  global target_g_table = [
  	"NaCl", "spatula_L", "6.5",
  	"NaCl", "spatula_M", "1.5",
  	"NaCl", "spatula_S", "0.135",

  	"Mannitol", "spatula_L", "2.85",
  	"Mannitol", "spatula_M", "0.8",
  	"Mannitol", "spatula_S", "0.075",

  	"CCS", "spatula_L", "2.45",
  	"CCS", "spatula_M", "0.6",
  	"CCS", "spatula_S", "0.075",

  	"lactose_loose", "spatula_L", "1.6",
  	"lactose_loose", "spatula_M", "0.5",
  	"lactose_loose", "spatula_S", "0.05",

  	"Magnesium_sterate", "spatula_flat_M", "0.6",
  	"Magnesium_sterate", "spatula_flat_S", "0.25",

  	"lactose_fine", "spatula_flat_M", "1.0",
  	"lactose_fine", "spatula_flat_S", "0.5"]

  def get_target_g(Pow_name, spat_name):
  	local i = 0
  	local n = length(target_g_table)
  	while (i < n):
  		if (target_g_table[i] == Pow_name and target_g_table[i+1] == spat_name):
  			return to_num(target_g_table[i+2])
  		end
  		i = i+3
  	end
  	popup("No target_g match for: ", Pow_name, ", ", spatula)

  end
  def auto_tilt_and_scoop(W_now, target_weight, Weight_value):
  	level = compute_level_percent(W_now, Weight_value)

  	#global angle_deg = compute_tilt_deg(level)

  	#if(level>=10.0):
  		#target_g = 2.850
  	#elif(level<10.0 and level >=1.0):
  		#target_g= 0.8
  	#else:
  		#target_g = 0.060
  	#end


  	#if (Task =="Emptying"):
  		#if (level>10.0):
  			#target_g = 2.850
  		#elif (level<=10.0 and level >1.0):
  			#target_g = 0.8
  		#else:
  			#target_g = 0.060
  		#end
  	#elif (Task == "Dosing"):
  		#if (level>10.0 and diff>=3.5):
  			#target_g = 2.85
  		#elif (level>10.0 and diff<3.5):
  			#target_g = 0.8
  		#elif (level<=10.0 and level >1.0):
  			#target_g = 0.8
  		#else:
  			#target_g = 0.06
  		#end
  	#end

  	global spatula = select_spatula(Pow_name, level, diff)
  	global target_g = get_target_g(Pow_name, spatula)

  	global scoop_depth = compute_scoop_depth(level, Weight_value, target_g)

  	tilt(level)
  	#P_center = get_actual_tcp_pose()

  	if (scoop_ct < 5 and g_prev_cum_w>0.0):
  		#local scoop_g = scoop_g
  		local error = target_g - scoop_g
  		error_sum = error_sum + error
  		error_sq_sum = error_sq_sum + error*error
  		scoop_ct = scoop_ct+1

  		if (scoop_ct==5):
  			local avg_error = error_sum/5.0
  			#local std_dev = sqrt(error_sq_sum/5.0) - (avg_error*avg_error))

  			if (my_abs(avg_error)>1.0):
  				g_k = 0.055
  				g_alpha = 0.85
  			elif (my_abs(avg_error)>0.6):
  				g_k= 0.045
  				g_alpha =0.75
  			elif (my_abs(avg_error)> 0.3):
  				g_k = 0.035
  				g_alpha = 0.65
  			elif (my_abs(avg_error)>0.1):
  				g_k = 0.025
  				g_alpha = 0.55
  			else:
  				g_k = 0.015
  				g_alpha = 0.45
  			end
  		end
  	end

  	scoop_powder(P_center)
  end


  def after_scoop():
  	tilt_send(angle_deg)
  	sleep(0.5)
  	movel(lifted_pose, a=0.05, v=0.2)
  	movel(tilted_pose_in_base, a=0.05, v=0.2)
  	set_analog_out(0,0.4)
  	movel(pose_trans(tilted_pose_in_base, p[-0.01,0,0,0,0,2.0]), a=0.05, v=0.2)
  	set_analog_out(0,0.0)
  	movel(lifted_pose, a=0.05, v=0.2)
  	tilt_to_home()
  end
  $ 23 "Script: Weight_scale_socket.script"
  def get_weight():
  	socket_open("192.168.12.190", 3002)
  	sleep(0.2)
  	textmsg("socket opened successfully!")
  	socket_send_string("GET_WEIGHT")
  	sync()
  	sleep(0.5)
  	receiveFromServ = socket_read_ascii_float(6)
  	while (receiveFromServ[0] <1):
  		sleep(0.5)
  		receiveFromServ = socket_read_ascii_float(1)
  		textmsg("retrying read:", receiveFromServ)
  	end
  	textmsg("Received weight:", receiveFromServ[1])
  	socket_close()
  	sleep(0.2)
  	return receiveFromServ[1]
  end

  def tare_scale():
  	socket_open("192.168.12.190", 3002)
  	socket_send_string("TARE")
  	sleep(0.5)
  	socket_close()
  end

  def zero_scale():
  	socket_open("192.168.12.190", 3002)
  	socket_send_string("ZERO")
  	sleep(0.5)
  	socket_close()
  end

  def log_weight():
  	socket_open("192.168.12.190", 3002)
  	socket_send_string("LOG_WEIGHT")
  	sleep(0.5)
  	socket_close()
  end
  $ 24 "BeforeStarts"
  $ 25 "uLM"
  $ 26 "CMD_Stop≔ False "
  global CMD_Stop=  False
  $ 27 "CMD_Abort≔ False "
  global CMD_Abort=  False
  $ 28 "CMD_Clear≔ False "
  global CMD_Clear=  False
  $ 29 "STATE≔1"
  global STATE=1
  $ 30 "STATE_Info≔''"
  global STATE_Info=""
  $ 31 "ARM_Referenced≔ False "
  global ARM_Referenced=  False
  $ 32 "zero_ftsensor()"
  zero_ftsensor()
  $ 33 "poses init"
  $ 34 "PSE_A≔p[0,0,0,0,0,0]"
  global PSE_A=p[0,0,0,0,0,0]
  $ 35 "PSE_A_H≔p[0,0,0,0,0,0]"
  global PSE_A_H=p[0,0,0,0,0,0]
  $ 36 "PSE_R≔p[0,0,0,0,0,0]"
  global PSE_R=p[0,0,0,0,0,0]
  $ 37 "PSE_R_H≔p[0,0,0,0,0,0]"
  global PSE_R_H=p[0,0,0,0,0,0]
  $ 38 "PSE_T≔p[0,0,0,0,0,0]"
  global PSE_T=p[0,0,0,0,0,0]
  $ 39 "PSE_T_H≔p[0,0,0,0,0,0]"
  global PSE_T_H=p[0,0,0,0,0,0]
  $ 40 "PSE_C_E≔p[0,0,0,0,0,0]"
  global PSE_C_E=p[0,0,0,0,0,0]
  $ 41 "PSE_C_H≔p[0,0,0,0,0,0]"
  global PSE_C_H=p[0,0,0,0,0,0]
  $ 42 "PSE_C_S≔p[0,0,0,0,0,0]"
  global PSE_C_S=p[0,0,0,0,0,0]
  $ 43 "init_home_by_cartesian_pose(p[0,-0.400,0.300,0,0,0])"
  init_home_by_cartesian_pose(p[0,-0.400,0.300,0,0,0])
  $ 44 "Clearing"
  $ 45 "reset_error()"
  reset_error()
  $ 46 "reset_warning()"
  reset_warning()
  $ 47 "uGo"
  $ 49 "ugo_init( True ,'http://192.168.12.120:10001')"
  ugo_init(  True  ,"http://192.168.12.120:10001")
  $ 50 "ugo_update_outputs()"
  ugo_update_outputs()
  $ 51 "App"
  $ 52 "'ADD APPLICATION SPECIFIC COMMANDS'"
  # 'ADD APPLICATION SPECIFIC COMMANDS'
  $ 53 "Tools"
  $ 54 "OBJ_Picked≔gripper_has_object()"
  global OBJ_Picked=gripper_has_object()
  $ 55 "If OBJ_Picked"
  if (OBJ_Picked):
    # begin: URCap Program Node
    #   Source: Robotiq_Grippers, 1.8.4.4844, Robotiq Inc.
    #   Type: Gripper Activate
    $ 56 "Gripper Activate"

    kill rq_gripper_communication_thread
    rq_gripper_communication_thread_started = False

    rq_init_comm_if_connected(9, "1")
    rq_init_comm_if_connected(2, "2")
    rq_init_comm_if_connected(3, "3")
    rq_init_comm_if_connected(4, "4")
    rq_print_connected_grippers()
    rq_gripper_communication_thread = run rq_gripper_communication()

    while(not rq_gripper_communication_thread_started):
        sync()
    end

    rq_set_max_current_for_all_grippers()

    reset_and_activate = False

    rq_activate_all_grippers(False)
    # end: URCap Program Node
  else:
    $ 57 "Else" "noBreak"
    # begin: URCap Program Node
    #   Source: Robotiq_Grippers, 1.8.4.4844, Robotiq Inc.
    #   Type: Gripper Activate
    $ 58 "Gripper Reset and Activate"

    kill rq_gripper_communication_thread
    rq_gripper_communication_thread_started = False

    rq_init_comm_if_connected(9, "1")
    rq_init_comm_if_connected(2, "2")
    rq_init_comm_if_connected(3, "3")
    rq_init_comm_if_connected(4, "4")
    rq_print_connected_grippers()
    rq_gripper_communication_thread = run rq_gripper_communication()

    while(not rq_gripper_communication_thread_started):
        sync()
    end

    rq_set_max_current_for_all_grippers()

    reset_and_activate = True

    rq_activate_all_grippers(True)
    # end: URCap Program Node
  end
  $ 59 "zero_ftsensor()"
  zero_ftsensor()
  $ 60 "EXTT"
  $ 61 "Set GRP_3F_Enable=Off"
  set_standard_digital_out(4, False)
  $ 62 "Set DO[6]=Off"
  set_standard_digital_out(6, False)
  $ 63 "Set GRP_3F_Decap=Off"
  set_standard_digital_out(3, False)
  $ 64 "Set GRP_3F_Cap=Off"
  set_standard_digital_out(2, False)
  $ 65 "Set GRP_3F_Open=Off"
  set_standard_digital_out(5, False)
  $ 66 "PSE_T≔get_tool_free_pose(dir=[0,0,0.150], move_in_base_frame=True)"
  global PSE_T=get_tool_free_pose(dir=[0,0,0.150], move_in_base_frame=True)
  $ 67 "If is_reachable(Base_const, [PSE_T])"
  if (is_reachable(p[0.0,0.0,0.0,0.0,0.0,0.0], [PSE_T])):
    $ 68 "MoveL"
    $ 69 "PSE_T" "breakAfter"
    movel(PSE_T, a=1.2, v=0.15)
  end
  $ 70 "powder dispensing variable init"
  $ 71 "Start_thread≔ False "
  global Start_thread=  False
  $ 72 "vib_mot_thread≔ False "
  global vib_mot_thread=  False
  $ 73 "kp≔0.0005"
  global kp=0.0005
  $ 74 "ki≔0.005"
  global ki=0.005
  $ 75 "kd≔0.02"
  global kd=0.02
  $ 76 "dt≔0.02"
  global dt=0.02
  $ 77 "Integral_error≔0"
  global Integral_error=0
  $ 78 "current_error≔0"
  global current_error=0
  $ 79 "previous_error≔0"
  global previous_error=0
  $ 80 "tilt_increment≔0"
  global tilt_increment=0
  $ 81 "tilt_angle≔0"
  global tilt_angle=0
  $ 82 "diff≔0"
  global diff=0
  $ 83 "current_pose≔get_actual_tcp_pose()"
  global current_pose= get_actual_tcp_pose ()
  $ 84 "Relative_trans≔p[0, 0, -0.035, 0, 0, 0]"
  global Relative_trans=p[0, 0, -0.035, 0, 0, 0]
  $ 85 "ContA_plc_offst≔p[-0.00205, 0.02547, 0.03730, -0.03, -2.183, 6.165]"
  global ContA_plc_offst=p[-0.00205, 0.02547, 0.03730, -0.03, -2.183, 6.165]
  $ 86 "PowA_50_offset≔p[0.21808, -0.19943, 0.06584, 0, 0, 0]"
  global PowA_50_offset=p[0.21808, -0.19943, 0.06584, 0, 0, 0]
  $ 88 "tilt_init_reference()"
  tilt_init_reference()
  $ 89 "switch_spat_M≔ True "
  global switch_spat_M=  True
  $ 90 "switch_spat_S≔ True "
  global switch_spat_S=  True
  $ 698 "Thread_1"
  thread Thread_1():
    while (True):
      $ 699 "If Start_thread≟ True "
      if (Start_thread ==   True  ):
        $ 700 "Weight_value≔get_weight()"
        global Weight_value=get_weight()
        $ 701 "Wait: 0.1"
        sleep(0.1)
        $ 702 "sync()"
        sync()
      end
    end
  end
  threadId_Thread_1 = run Thread_1()
  while (True):
    $ 91 "Robot Program"
    $ 92 "MAIN"
    $ 93 "command_manager(external_control='uGO', cond_suspend=(ITM_Manipulated and AMR_AtTarget and AMR_Charging and AMR_Battery<40), cond_unsuspend=(AMR_Battery≟60))"
    command_manager(external_control="uGO", cond_suspend=(ITM_Manipulated  and  AMR_AtTarget  and  AMR_Charging  and  AMR_Battery<40), cond_unsuspend=(AMR_Battery == 60))
    $ 94 "log_state(STATE_Info)"
    log_state(STATE_Info)
    $ 95 "Switch STATE"
    switch_1 = STATE
    $ 96 "Case 1"
    if (1 == switch_1):
      $ 97 "Stopping"
      $ 98 "STATE_Info≔'Stopping'"
      global STATE_Info="Stopping"
      $ 99 "end_freedrive_mode()"
      end_freedrive_mode()
      $ 100 "Set"
      set_tcp(p[0.0,0.0,0.161,3.1415,0.0,0.0])
      $ 101 "PSE_T≔get_tool_free_pose(dir=[0,0,0.150], move_in_base_frame=True)"
      global PSE_T=get_tool_free_pose(dir=[0,0,0.150], move_in_base_frame=True)
      $ 102 "If is_reachable(Base_const, [PSE_T])"
      if (is_reachable(p[0.0,0.0,0.0,0.0,0.0,0.0], [PSE_T])):
        $ 103 "MoveL"
        $ 104 "PSE_T" "breakAfter"
        movel(PSE_T, a=1.2, v=0.15)
      end
      $ 105 "do_transition(keep_rxry=OBJ_Picked, r=0)"
      do_transition(keep_rxry=OBJ_Picked, r=0)
      $ 115 "If stopping() and AMR_Done"
      if (stopping()  and  AMR_Done):
        $ 116 "STATE≔2"
        global STATE=2
        $ 117 "ugo_update_outputs()"
        ugo_update_outputs()
      end
    elif (2 == switch_1):
      $ 118 "Case 2"
      $ 119 "Stopped"
      $ 120 "STATE_Info≔'Stopped'"
      global STATE_Info="Stopped"
      $ 122 "If CMD_Reset"
      if (CMD_Reset):
        $ 123 "STATE≔3"
        global STATE=3
        $ 124 "ugo_update_outputs()"
        ugo_update_outputs()
      end
    elif (3 == switch_1):
      $ 125 "Case 3"
      $ 126 " Resetting"
      $ 127 "STATE_Info≔'Resetting'"
      global STATE_Info="Resetting"
      $ 128 "uML"
      $ 129 "reset_error()"
      reset_error()
      $ 130 "reset_warning()"
      reset_warning()
      $ 131 "PROCESS_Step≔0"
      global PROCESS_Step=0
      $ 132 "PROCESS_Info≔''"
      global PROCESS_Info=""
      $ 133 "ARM_Referenced≔ False "
      global ARM_Referenced=  False
      $ 134 "WRK_Done≔ False "
      global WRK_Done=  False
      $ 135 "ITM_Prepared≔ False "
      global ITM_Prepared=  False
      $ 136 "ITM_Manipulated≔ False "
      global ITM_Manipulated=  False
      $ 137 "STP≔0"
      global STP=0
      $ 138 "Action≔0"
      global Action=0
      $ 139 "Action_Info≔''"
      global Action_Info=""
      $ 140 "ITM_ID≔0"
      global ITM_ID=0
      $ 141 "JIG≔0"
      global JIG=0
      $ 142 "JIG_Slot≔0"
      global JIG_Slot=0
      $ 143 "Task_info≔''"
      global Task_info=""
      $ 144 "Set"
      set_tcp(p[0.0,0.0,0.161,3.1415,0.0,0.0])
      $ 145 "App"
      $ 146 "'ADD APPLICATION SPECIFIC COMMANDS'"
      # 'ADD APPLICATION SPECIFIC COMMANDS'
      $ 147 "OBJ_Type≔0"
      global OBJ_Type=0
      $ 148 "OBJ_Nbr≔0"
      global OBJ_Nbr=0
      $ 149 "If CNT_Rack_Output≥50"
      if (CNT_Rack_Output >= 50):
        $ 150 "CNT_Rack_Output≔0"
        global CNT_Rack_Output=0
      end
      $ 151 "TASK≔struct(ID=0, NAVI=struct(target=0, footprint=0, protectiveOff=0, dock=0), WORK=struct(ITM_ID_Src=0, JIG_ID_Src=0, OBJ_Nbr_Src=0, ACT_Src=0, ITM_ID_Tgt=0, JIG_ID_Tgt=0, OBJ_Nbr_Tgt=0, ACT_Tgt=0, OBJ_Type=0))"
      global TASK=struct(ID=0, NAVI=struct(target=0, footprint=0, protectiveOff=0, dock=0), WORK=struct(ITM_ID_Src=0, JIG_ID_Src=0, OBJ_Nbr_Src=0, ACT_Src=0, ITM_ID_Tgt=0, JIG_ID_Tgt=0, OBJ_Nbr_Tgt=0, ACT_Tgt=0, OBJ_Type=0))
      $ 153 "If resetting() and AMR_Done"
      if (resetting()  and  AMR_Done):
        $ 154 "STATE≔4"
        global STATE=4
        $ 155 "ugo_update_outputs()"
        ugo_update_outputs()
      end
    elif (4 == switch_1):
      $ 156 "Case 4"
      $ 157 "Idle"
      $ 158 "STATE_Info≔'Idle'"
      global STATE_Info="Idle"
      $ 159 "If CMD_Start"
      if (CMD_Start):
        $ 160 "STATE≔5"
        global STATE=5
        $ 161 "ugo_update_outputs()"
        ugo_update_outputs()
      end
    elif (5 == switch_1):
      $ 162 "Case 5"
      $ 163 "Starting"
      $ 164 "STATE_Info≔'Starting'"
      global STATE_Info="Starting"
      $ 165 "'ADD COMMANDS WHAT TO START WITH'"
      # 'ADD COMMANDS WHAT TO START WITH'
      $ 167 "get ugo data"
      $ 168 "Assign Tasks"
      $ 169 "TASK.ID = ugo_get_task()"
      TASK.ID = ugo_get_task()
      $ 170 "If TASK.ID≟1"
      if (TASK.ID == 1):
        $ 171 "Task_info≔'Charge'"
        global Task_info="Charge"
        $ 172 "Parameters"
        $ 173 "AMR_PosTarget≔1"
        global AMR_PosTarget=1
      else:
        $ 174 "ElseIf TASK.ID≟9"
        if (TASK.ID == 9):
          $ 175 "'Pick Sarstedt Rack from Variable source'"
          # 'Pick Sarstedt Rack from Variable source'
          $ 176 "Task_info≔'Navigate to Target'"
          global Task_info="Navigate to Target"
          $ 177 "Parameters"
          $ 178 "AMR_PosTarget≔UGO.read_input('00','ITM_ID')"
          global AMR_PosTarget=UGO.read_input("00","ITM_ID")
        else:
          $ 179 "ElseIf TASK.ID≟49"
          if (TASK.ID == 49):
            $ 180 "Task_info≔'Pick Containers'"
            global Task_info="Pick Containers"
            $ 181 "Parameters"
            $ 182 "ITM_ID≔1"
            global ITM_ID=1
            $ 183 "OBJ_Type≔6"
            global OBJ_Type=6
            $ 184 "JIG≔15"
            global JIG=15
            $ 185 "AMR_PosTarget≔3"
            global AMR_PosTarget=3
          else:
            $ 186 "ElseIf TASK.ID≟50"
            if (TASK.ID == 50):
              $ 187 "Task_info≔'Decap Containers'"
              global Task_info="Decap Containers"
              $ 188 "Parameters"
              $ 189 "ITM_ID≔1"
              global ITM_ID=1
              $ 190 "OBJ_Type≔6"
              global OBJ_Type=6
              $ 191 "JIG≔16"
              global JIG=16
              $ 192 "AMR_PosTarget≔5"
              global AMR_PosTarget=5
            else:
              $ 193 "ElseIf TASK.ID≟51"
              if (TASK.ID == 51):
                $ 194 "Task_info≔'Detect Spatula and transfer powder'"
                global Task_info="Detect Spatula and transfer powder"
                $ 195 "Parameters"
                $ 196 "ITM_ID≔1"
                global ITM_ID=1
                $ 197 "Target_weight≔(UGO.read_input('00','Target_weight'))/1000"
                global Target_weight=(UGO.read_input("00","Target_weight"))/1000
                $ 198 "OBJ_Type≔8"
                global OBJ_Type=8
                $ 199 "JIG≔16"
                global JIG=16
                $ 200 "AMR_PosTarget≔5"
                global AMR_PosTarget=5
              else:
                $ 201 "ElseIf TASK.ID≟52"
                if (TASK.ID == 52):
                  $ 202 "Task_info≔'Pick PowderA'"
                  global Task_info="Pick PowderA"
                  $ 203 "Parameters"
                  $ 204 "ITM_ID≔1"
                  global ITM_ID=1
                  $ 205 "OBJ_Type≔6"
                  global OBJ_Type=6
                  $ 206 "JIG≔15"
                  global JIG=15
                  $ 207 "AMR_PosTarget≔3"
                  global AMR_PosTarget=3
                else:
                  $ 208 "ElseIf TASK.ID≟53"
                  if (TASK.ID == 53):
                    $ 209 "Task_info≔'Decap PowderA'"
                    global Task_info="Decap PowderA"
                    $ 210 "Parameters"
                    $ 211 "ITM_ID≔1"
                    global ITM_ID=1
                    $ 212 "OBJ_Type≔6"
                    global OBJ_Type=6
                    $ 213 "JIG≔1"
                    global JIG=1
                    $ 214 "AMR_PosTarget≔5"
                    global AMR_PosTarget=5
                  else:
                    $ 215 "ElseIf TASK.ID≟54"
                    if (TASK.ID == 54):
                      $ 216 "Task_info≔'Empty PowderA'"
                      global Task_info="Empty PowderA"
                      $ 217 "Parameters"
                      $ 218 "ITM_ID≔1"
                      global ITM_ID=1
                      $ 219 "Target_weight≔(UGO.read_input('00','Target_weight'))/1000"
                      global Target_weight=(UGO.read_input("00","Target_weight"))/1000
                      $ 220 "W_now≔(UGO.read_input('00','Container_weight'))/1000"
                      global W_now=(UGO.read_input("00","Container_weight"))/1000
                      $ 221 "Powder_name≔(UGO.read_input('00','Powder_name'))"
                      global Powder_name=(UGO.read_input("00","Powder_name"))
                      $ 222 "OBJ_Type≔6"
                      global OBJ_Type=6
                      $ 223 "JIG≔17"
                      global JIG=17
                      $ 224 "AMR_PosTarget≔5"
                      global AMR_PosTarget=5
                    else:
                      $ 225 "ElseIf TASK.ID≟55"
                      if (TASK.ID == 55):
                        $ 226 "Task_info≔'Place PowderA'"
                        global Task_info="Place PowderA"
                        $ 227 "Parameters"
                        $ 228 "ITM_ID≔1"
                        global ITM_ID=1
                        $ 229 "OBJ_Type≔6"
                        global OBJ_Type=6
                        $ 230 "JIG≔21"
                        global JIG=21
                        $ 231 "AMR_PosTarget≔5"
                        global AMR_PosTarget=5
                      else:
                        $ 232 "ElseIf TASK.ID≟56"
                        if (TASK.ID == 56):
                          $ 233 "Task_info≔'Dose Powder'"
                          global Task_info="Dose Powder"
                          $ 234 "Parameters"
                          $ 235 "ITM_ID≔1"
                          global ITM_ID=1
                          $ 236 "Target_weight≔(UGO.read_input('00','Target_weight'))/1000"
                          global Target_weight=(UGO.read_input("00","Target_weight"))/1000
                          $ 237 "W_now≔(UGO.read_input('00','Container_weight'))/1000"
                          global W_now=(UGO.read_input("00","Container_weight"))/1000
                          $ 238 "Pow_name≔(UGO.read_input('00','Powder_name'))"
                          global Pow_name=(UGO.read_input("00","Powder_name"))
                          $ 239 "OBJ_Type≔6"
                          global OBJ_Type=6
                          $ 240 "JIG≔17"
                          global JIG=17
                          $ 241 "AMR_PosTarget≔5"
                          global AMR_PosTarget=5
                        else:
                          $ 242 "Else" "noBreak"
                          $ 243 "set_error(ERROR_WRONG_ORDER)"
                          set_error(ERROR_WRONG_ORDER)
                        end
                      end
                    end
                  end
                end
              end
            end
          end
        end
      end
      $ 244 "test ugo"
      $ 245 "Wait: 0.2"
      sleep(0.2)
      $ 246 "ugo_update_outputs()"
      ugo_update_outputs()
      $ 247 "If starting() and AMR_Done"
      if (starting()  and  AMR_Done):
        $ 248 "log_message(Task_info, 'New Task: ')"
        log_message(Task_info, "New Task: ")
        $ 249 "log_message(to_str(TASK.ID), 'Task_ID: ')"
        log_message(to_str(TASK.ID), "Task_ID: ")
        $ 250 "do_transition(keep_rxry=OBJ_Picked)"
        do_transition(keep_rxry=OBJ_Picked)
        $ 251 "STATE≔6"
        global STATE=6
        $ 252 "ugo_update_outputs()"
        ugo_update_outputs()
      end
    elif (6 == switch_1):
      $ 253 "Case 6"
      $ 254 "Execute"
      $ 255 "STATE_Info≔'Execute'"
      global STATE_Info="Execute"
      $ 256 "If  not CMD_Hold and not CMD_Suspend"
      global thread_flag_256=0
      thread Thread_if_256():
        $ 257 "Switch PROCESS_Step"
        switch_2 = PROCESS_Step
        $ 258 "Case 0"
        if (0 == switch_2):
          $ 259 "PROCESS_Info≔'process control'"
          global PROCESS_Info="process control"
          $ 260 "log_process(PROCESS_Info)"
          log_process(PROCESS_Info)
          $ 261 "process control"
          $ 262 "If  not AMR_AtTarget"
          if (  not  AMR_AtTarget):
            $ 263 "PROCESS_Step≔1"
            global PROCESS_Step=1
          else:
            $ 264 "ElseIf (( not ITM_Prepared and  not WRK_Done) or (ITM_Prepared and WRK_Done))"
            if (((  not  ITM_Prepared  and    not  WRK_Done)  or  (ITM_Prepared  and  WRK_Done))):
              $ 265 "PROCESS_Step≔2"
              global PROCESS_Step=2
            else:
              $ 266 "ElseIf  not WRK_Done"
              if (  not  WRK_Done):
                $ 267 "PROCESS_Step≔3"
                global PROCESS_Step=3
              else:
                $ 268 "Else" "noBreak"
                $ 269 "task finished"
                $ 270 "PROCESS_Info≔''"
                global PROCESS_Info=""
                $ 271 "STATE≔7"
                global STATE=7
                $ 272 "ugo_update_outputs()"
                ugo_update_outputs()
              end
            end
          end
        elif (1 == switch_2):
          $ 273 "Case 1"
          $ 274 "navigate"
          $ 275 "'MOVING THE uML'"
          # 'MOVING THE uML'
          $ 276 "PROCESS_Info≔'move to target'"
          global PROCESS_Info="move to target"
          $ 277 "log_process(PROCESS_Info)"
          log_process(PROCESS_Info)
          $ 278 "If TASK.ID≟1"
          if (TASK.ID == 1):
            $ 279 "Action≔51"
            global Action=51
          else:
            $ 280 "Else" "noBreak"
            $ 281 "Action≔52"
            global Action=52
          end
          $ 283 "If AMR_Done"
          if (AMR_Done):
            $ 284 "PROCESS_Step≔0"
            global PROCESS_Step=0
          end
        elif (2 == switch_2):
          $ 285 "Case 2"
          $ 286 "prepare"
          $ 287 "'THINGS THAT HAVE TO BE DONE ONCE IN A SEQUENCE,WORKFLOW'"
          # 'THINGS THAT HAVE TO BE DONE ONCE IN A SEQUENCE,WORKFLOW'
          $ 288 "PROCESS_Info≔'prepare for work'"
          global PROCESS_Info="prepare for work"
          $ 289 "log_process(PROCESS_Info)"
          log_process(PROCESS_Info)
          $ 290 "If TASK.WORK.ITM_ID_Src>1"
          if (TASK.WORK.ITM_ID_Src>1):
            $ 291 "ITM_ID≔TASK.WORK.ITM_ID_Src"
            global ITM_ID=TASK.WORK.ITM_ID_Src
          else:
            $ 292 "ElseIf TASK.WORK.ITM_ID_Tgt>1"
            if (TASK.WORK.ITM_ID_Tgt>1):
              $ 293 "ITM_ID≔TASK.WORK.ITM_ID_Tgt"
              global ITM_ID=TASK.WORK.ITM_ID_Tgt
            end
          end
          $ 294 "If  not ARM_Referenced and (ITM_ID≠0)"
          if (  not  ARM_Referenced  and  (ITM_ID != 0)):
            $ 295 "STP≔1"
            global STP=1
          else:
            $ 296 "ElseIf ARM_Referenced or (ITM_ID≟0)"
            if (ARM_Referenced  or  (ITM_ID == 0)):
              $ 297 "STP≔2"
              global STP=2
            end
          end
          $ 298 "Switch STP"
          switch_3 = STP
          $ 299 "Case 1"
          if (1 == switch_3):
            $ 300 "reference"
            $ 301 "STP_Info≔'reference at target position'"
            global STP_Info="reference at target position"
            $ 302 "log_step(STP_Info)"
            log_step(STP_Info)
            $ 303 "If ITM_ID≟1"
            if (ITM_ID == 1):
              $ 304 "CAM_Done≔ True "
              global CAM_Done=  True
            else:
              $ 305 "Else" "noBreak"
              $ 306 "Action≔131"
              global Action=131
              $ 307 "Call Sub_Vision_V18"
              Sub_Vision_V18()
            end
            $ 309 "If CAM_Done and  not ERROR.FLAG"
            if (CAM_Done  and    not  ERROR.FLAG):
              $ 310 "log_step('ARM referenced')"
              log_step("ARM referenced")
              $ 311 "ARM_Referenced≔ True "
              global ARM_Referenced=  True
            end
          elif (2 == switch_3):
            $ 312 "Case 2"
            $ 313 "manipulate"
            $ 314 "STP_Info≔'manipulate item'"
            global STP_Info="manipulate item"
            $ 315 "log_step(STP_Info)"
            log_step(STP_Info)
            $ 316 "'In case pressing button is needed'"
            # 'In case pressing button is needed'
            $ 317 "If found_in_list(ITM_ID, ITM_ID_List)"
            if (found_in_list(ITM_ID, ITM_ID_List)):
              $ 318 "Switch ITM_ID"
              switch_4 = ITM_ID
              $ 319 "Case 0"
              if (0 == switch_4):
                $ 320 "ITM_Manipulated≔ not ITM_Manipulated"
                global ITM_Manipulated=  not  ITM_Manipulated
              elif (1 == switch_4):
                $ 321 "Case 1"
                $ 322 "ITM_Manipulated≔ not ITM_Manipulated"
                global ITM_Manipulated=  not  ITM_Manipulated
              elif (2 == switch_4):
                $ 323 "Case 2"
              else:
                $ 333 "Default Case"
                $ 334 "ITM_Manipulated≔ not ITM_Manipulated"
                global ITM_Manipulated=  not  ITM_Manipulated
              end
            end
          end
          $ 335 "ITM_Prepared≔(ITM_Manipulated or  not found_in_list(ITM_ID, ITM_ID_List)) and (ARM_Referenced or ITM_ID≟0) and  not WRK_Done"
          global ITM_Prepared=(ITM_Manipulated  or    not  found_in_list(ITM_ID, ITM_ID_List))  and  (ARM_Referenced  or  ITM_ID == 0)  and    not  WRK_Done
          $ 336 "STP≔0"
          global STP=0
          $ 337 "STP_Info≔''"
          global STP_Info=""
          $ 338 "PROCESS_Step≔0"
          global PROCESS_Step=0
        elif (3 == switch_2):
          $ 339 "Case 3"
          $ 340 "work"
          $ 341 "'ADD EVERY MACHINE, OBJECT, STATION TO WORK ON'"
          # 'ADD EVERY MACHINE, OBJECT, STATION TO WORK ON'
          $ 342 "Switch ITM_ID"
          switch_3 = ITM_ID
          $ 343 "Case 1"
          if (1 == switch_3):
            $ 344 "uLM"
            $ 345 "If TASK.ID≟12"
            if (TASK.ID == 12):
              $ 346 "fill racks"
              $ 347 "Action≔151"
              global Action=151
              $ 348 "Call Sub_Vision_V18"
              Sub_Vision_V18()
              $ 349 "If  not ERROR.FLAG"
              if (  not  ERROR.FLAG):
                $ 350 "Actions for the task"
                $ 351 "Action≔1"
                global Action=1
                $ 352 "JIG≔2"
                global JIG=2
                $ 353 "JIG_Slot≔CAM_Result[0]"
                global JIG_Slot=CAM_Result[0]
                $ 354 "OBJ_Nbr≔CAM_Result[0]"
                global OBJ_Nbr=CAM_Result[0]
                $ 355 "OBJ_Type≔2"
                global OBJ_Type=2
                $ 356 "Call Sub_Action_V4"
                Sub_Action_V4()
                $ 357 "If OBJ_Picked"
                if (OBJ_Picked):
                  $ 358 "CAM_Result.remove(0)"
                  CAM_Result.remove(0)
                  $ 359 "PRC_TubCounter≔PRC_TubCounter+1"
                  global PRC_TubCounter=PRC_TubCounter+1
                  $ 360 "If PRC_TubCounter%4≟0"
                  if (PRC_TubCounter%4 == 0):
                    $ 361 "JIG_Slot≔4"
                    global JIG_Slot=4
                  else:
                    $ 362 "Else" "noBreak"
                    $ 363 "JIG_Slot≔PRC_TubCounter%4"
                    global JIG_Slot=PRC_TubCounter%4
                  end
                  $ 364 "OBJ_Nbr≔ceil(PRC_TubCounter/4)"
                  global OBJ_Nbr=ceil(PRC_TubCounter/4)
                  $ 365 "Action≔2"
                  global Action=2
                  $ 366 "JIG≔4"
                  global JIG=4
                  $ 367 "Call Sub_Action_V4"
                  Sub_Action_V4()
                  $ 368 "Action≔151"
                  global Action=151
                  $ 369 "Call Sub_Vision_V18"
                  Sub_Vision_V18()
                end
              end
              $ 370 "If (CAM_Captures≥CAM_PRM_Retries) or (PRC_TubCounter≥32)"
              if ((CAM_Captures >= CAM_PRM_Retries)  or  (PRC_TubCounter >= 32)):
                $ 371 "PROCESS_Step≔0"
                global PROCESS_Step=0
                $ 372 "WRK_Done≔ True "
                global WRK_Done=  True
              end
            else:
              $ 373 "ElseIf TASK.ID≟49"
              if (TASK.ID == 49):
                $ 374 "Pick Powder container"
                $ 375 "Action≔131"
                global Action=131
                $ 376 "Call Sub_Vision_V18"
                Sub_Vision_V18()
                $ 377 "Action≔35"
                global Action=35
                $ 378 "Call Sub_Action_V4"
                Sub_Action_V4()
                $ 379 "PROCESS_Step≔0"
                global PROCESS_Step=0
                $ 380 "WRK_Done≔ True "
                global WRK_Done=  True
              else:
                $ 381 "ElseIf TASK.ID≟50"
                if (TASK.ID == 50):
                  $ 382 "Decap containers"
                  $ 383 "Action≔36"
                  global Action=36
                  $ 384 "Call Sub_Action_V4"
                  Sub_Action_V4()
                  $ 385 "PROCESS_Step≔0"
                  global PROCESS_Step=0
                  $ 386 "WRK_Done≔ True "
                  global WRK_Done=  True
                else:
                  $ 387 "ElseIf TASK.ID≟51"
                  if (TASK.ID == 51):
                    $ 388 "Detect Spatula and transfer powder"
                    $ 389 "Action≔131"
                    global Action=131
                    $ 390 "Call Sub_Vision_V18"
                    Sub_Vision_V18()
                    $ 391 "Action≔37"
                    global Action=37
                    $ 392 "Call Sub_Action_V4"
                    Sub_Action_V4()
                    $ 393 "PROCESS_Step≔0"
                    global PROCESS_Step=0
                    $ 394 "WRK_Done≔ True "
                    global WRK_Done=  True
                  else:
                    $ 395 "ElseIf TASK.ID≟52"
                    if (TASK.ID == 52):
                      $ 396 "Pick PowderA container"
                      $ 397 "Action≔131"
                      global Action=131
                      $ 398 "Call Sub_Vision_V18"
                      Sub_Vision_V18()
                      $ 399 "Action≔38"
                      global Action=38
                      $ 400 "Call Sub_Action_V4"
                      Sub_Action_V4()
                      $ 401 "PROCESS_Step≔0"
                      global PROCESS_Step=0
                      $ 402 "WRK_Done≔ True "
                      global WRK_Done=  True
                    else:
                      $ 403 "ElseIf TASK.ID≟53"
                      if (TASK.ID == 53):
                        $ 404 "Decap containerA"
                        $ 405 "Action≔39"
                        global Action=39
                        $ 406 "Call Sub_Action_V4"
                        Sub_Action_V4()
                        $ 407 "PROCESS_Step≔0"
                        global PROCESS_Step=0
                        $ 408 "WRK_Done≔ True "
                        global WRK_Done=  True
                      else:
                        $ 409 "ElseIf TASK.ID≟55"
                        if (TASK.ID == 55):
                          $ 410 "Place Powder"
                          $ 411 "Action≔131"
                          global Action=131
                          $ 412 "Call Sub_Vision_V18"
                          Sub_Vision_V18()
                          $ 413 "Action≔40"
                          global Action=40
                          $ 414 "Call Sub_Action_V4"
                          Sub_Action_V4()
                          $ 415 "PROCESS_Step≔0"
                          global PROCESS_Step=0
                          $ 416 "WRK_Done≔ True "
                          global WRK_Done=  True
                        else:
                          $ 417 "ElseIf TASK.ID≟54"
                          if (TASK.ID == 54):
                            $ 418 "Dispense Powder to Empty"
                            $ 419 "Action≔131"
                            global Action=131
                            $ 420 "Call Sub_Vision_V18"
                            Sub_Vision_V18()
                            $ 421 "Action≔41"
                            global Action=41
                            $ 422 "Call Sub_Action_V4"
                            Sub_Action_V4()
                            $ 423 "PROCESS_Step≔0"
                            global PROCESS_Step=0
                            $ 424 "WRK_Done≔ True "
                            global WRK_Done=  True
                          else:
                            $ 425 "ElseIf TASK.ID≟56"
                            if (TASK.ID == 56):
                              $ 426 "Dispense Powder"
                              $ 427 "Action≔131"
                              global Action=131
                              $ 428 "Call Sub_Vision_V18"
                              Sub_Vision_V18()
                              $ 429 "Action≔42"
                              global Action=42
                              $ 430 "Call Sub_Action_V4"
                              Sub_Action_V4()
                              $ 431 "PROCESS_Step≔0"
                              global PROCESS_Step=0
                              $ 432 "WRK_Done≔ True "
                              global WRK_Done=  True
                            end
                          end
                        end
                      end
                    end
                  end
                end
              end
            end
          elif (2 == switch_3):
            $ 433 "Case 2"
          elif (5 == switch_3):
            $ 475 "Case 5"
          elif (20 == switch_3):
            $ 483 "Case 20"
          elif (43 == switch_3):
            $ 545 "Case 43"
          else:
            $ 553 "Default Case"
            $ 554 "WRK_Done≔ True "
            global WRK_Done=  True
            $ 555 "PROCESS_Step≔0"
            global PROCESS_Step=0
          end
        end
        thread_flag_256 = 1
      end
      if (  not  CMD_Hold and not CMD_Suspend):
        global thread_handler_256=run Thread_if_256()
        while (thread_flag_256 == 0):
          if not(  not  CMD_Hold and not CMD_Suspend):
            kill thread_handler_256
            thread_flag_256 = 2
          else:
            sync()
          end
        end
      else:
        thread_flag_256 = 2
      end
      $ 556 "If CMD_Hold"
      if (CMD_Hold):
        $ 557 "STATE≔9"
        global STATE=9
        $ 558 "ugo_update_outputs()"
        ugo_update_outputs()
      else:
        $ 559 "ElseIf CMD_Suspend"
        if (CMD_Suspend):
          $ 560 "STATE≔12"
          global STATE=12
          $ 561 "ugo_update_outputs()"
          ugo_update_outputs()
        end
      end
    elif (7 == switch_1):
      $ 562 "Case 7"
      $ 563 "Completing"
      $ 564 "STATE_Info≔'Completing'"
      global STATE_Info="Completing"
      $ 565 "'ADD COMMANDS FOR COMPLETING THE PROCESS'"
      # 'ADD COMMANDS FOR COMPLETING THE PROCESS'
      $ 566 "do_transition(keep_rxry=OBJ_Picked)"
      do_transition(keep_rxry=OBJ_Picked)
      $ 568 "If completing() and AMR_Done"
      if (completing()  and  AMR_Done):
        $ 569 "STATE≔8"
        global STATE=8
        $ 570 "ugo_update_outputs()"
        ugo_update_outputs()
      end
    elif (8 == switch_1):
      $ 571 "Case 8"
      $ 572 "Complete"
      $ 573 "STATE_Info≔'Complete'"
      global STATE_Info="Complete"
      $ 574 "If CMD_Reset"
      if (CMD_Reset):
        $ 575 "STATE≔3"
        global STATE=3
        $ 576 "ugo_update_outputs()"
        ugo_update_outputs()
      end
    elif (9 == switch_1):
      $ 577 "Case 9"
      $ 578 "Holding"
      $ 579 "STATE_Info≔'Holding'"
      global STATE_Info="Holding"
      $ 580 "stopl(0.5)"
      stopl(0.5)
      $ 582 "If holding() and AMR_Done"
      if (holding()  and  AMR_Done):
        $ 583 "STATE≔10"
        global STATE=10
        $ 584 "ugo_update_outputs()"
        ugo_update_outputs()
      end
    elif (10 == switch_1):
      $ 585 "Case 10"
      $ 586 "Held"
      $ 587 "STATE_Info≔'Held'"
      global STATE_Info="Held"
      $ 588 "If CMD_Unhold"
      if (CMD_Unhold):
        $ 589 "end_freedrive_mode()"
        end_freedrive_mode()
        $ 590 "STATE≔11"
        global STATE=11
        $ 591 "ugo_update_outputs()"
        ugo_update_outputs()
      else:
        $ 592 "ElseIf FNC_Freedrive"
        if (FNC_Freedrive):
          $ 593 "freedrive_mode()"
          freedrive_mode()
        else:
          $ 594 "Else" "noBreak"
          $ 595 "end_freedrive_mode()"
          end_freedrive_mode()
        end
      end
    elif (11 == switch_1):
      $ 596 "Case 11"
      $ 597 "Unholding"
      $ 598 "STATE_Info≔'Unholding'"
      global STATE_Info="Unholding"
      $ 599 "Clearing"
      $ 600 "Switch ERROR.ID"
      switch_2 = ERROR.ID
      $ 601 "Case 1002"
      if (1002 == switch_2):
        $ 602 "AMR_AtTarget≔ False "
        global AMR_AtTarget=  False
        $ 603 "ARM_Referenced≔ False "
        global ARM_Referenced=  False
        $ 604 "ITM_Prepared≔ False "
        global ITM_Prepared=  False
        $ 605 "PROCESS_Step≔1"
        global PROCESS_Step=1
      elif (2007 == switch_2):
        $ 606 "Case 2007"
        $ 607 "PROCESS_Step≔1"
        global PROCESS_Step=1
      end
      $ 608 "reset_error()"
      reset_error()
      $ 609 "reset_warning()"
      reset_warning()
      $ 610 "OBJ_Picked≔gripper_has_object()"
      global OBJ_Picked=gripper_has_object()
      $ 612 "If unholding() and AMR_Done"
      if (unholding()  and  AMR_Done):
        $ 613 "STATE≔6"
        global STATE=6
        $ 614 "ugo_update_outputs()"
        ugo_update_outputs()
      end
    elif (12 == switch_1):
      $ 615 "Case 12"
      $ 616 "Suspending"
      $ 617 "STATE_Info≔'Suspending'"
      global STATE_Info="Suspending"
      $ 618 "PROCESS_Info≔str_cat(PROCESS_Info, ' suspended')"
      global PROCESS_Info=str_cat(PROCESS_Info, " suspended")
      $ 619 "If suspending()"
      if (suspending()):
        $ 620 "STATE≔13"
        global STATE=13
        $ 621 "ugo_update_outputs()"
        ugo_update_outputs()
      end
    elif (13 == switch_1):
      $ 622 "Case 13"
      $ 623 "Suspended"
      $ 624 "STATE_Info≔'Suspended'"
      global STATE_Info="Suspended"
      $ 626 "If CMD_Unsuspend"
      if (CMD_Unsuspend):
        $ 627 "STATE≔14"
        global STATE=14
        $ 628 "ugo_update_outputs()"
        ugo_update_outputs()
      end
    elif (14 == switch_1):
      $ 629 "Case 14"
      $ 630 "Unsuspending"
      $ 631 "STATE_Info≔'Unsuspending'"
      global STATE_Info="Unsuspending"
      $ 632 "PROCESS_Step≔0"
      global PROCESS_Step=0
      $ 633 "If unsuspending()"
      if (unsuspending()):
        $ 634 "STATE≔6"
        global STATE=6
        $ 635 "ugo_update_outputs()"
        ugo_update_outputs()
      end
    elif (15 == switch_1):
      $ 636 "Case 15"
      $ 637 "Aborting"
      $ 638 "STATE_Info≔'Aborting'"
      global STATE_Info="Aborting"
      $ 639 "If aborting()"
      if (aborting()):
        $ 640 "STATE≔16"
        global STATE=16
        $ 641 "ugo_update_outputs()"
        ugo_update_outputs()
      end
    elif (16 == switch_1):
      $ 642 "Case 16"
      $ 643 "Aborted"
      $ 644 "STATE_Info≔'Aborted'"
      global STATE_Info="Aborted"
      $ 645 "If CMD_Clear"
      if (CMD_Clear):
        $ 646 "STATE≔17"
        global STATE=17
        $ 647 "ugo_update_outputs()"
        ugo_update_outputs()
      end
    elif (17 == switch_1):
      $ 648 "Case 17"
      $ 649 "Clearing"
      $ 650 "STATE_Info≔'Clearing'"
      global STATE_Info="Clearing"
      $ 651 "Clearing"
      $ 652 "reset_warning()"
      reset_warning()
      $ 653 "reset_error()"
      reset_error()
      $ 654 "If clearing()"
      if (clearing()):
        $ 655 "STATE≔2"
        global STATE=2
        $ 656 "ugo_update_outputs()"
        ugo_update_outputs()
      end
    end
    $ 657 "log_state(STATE_Info)"
    log_state(STATE_Info)
    $ 658 "log_warning(WARNING.MSG)"
    log_warning(WARNING.MSG)
    $ 659 "log_error(ERROR.MSG)"
    log_error(ERROR.MSG)
    $ 660 "Times"
    $ 661 "Switch STATE"
    switch_1 = STATE
    $ 662 "Case 1"
    if (1 == switch_1):
      $ 663 "TM_St_Stopping≔get_time(STATE_Times[STATE-1])"
      global TM_St_Stopping=get_time(STATE_Times[STATE-1])
    elif (2 == switch_1):
      $ 664 "Case 2"
      $ 665 "TM_St_Stopped≔get_time(STATE_Times[STATE-1])"
      global TM_St_Stopped=get_time(STATE_Times[STATE-1])
    elif (3 == switch_1):
      $ 666 "Case 3"
      $ 667 "TM_St_Resetting≔get_time(STATE_Times[STATE-1])"
      global TM_St_Resetting=get_time(STATE_Times[STATE-1])
    elif (4 == switch_1):
      $ 668 "Case 4"
      $ 669 "TM_St_Idle≔get_time(STATE_Times[STATE-1])"
      global TM_St_Idle=get_time(STATE_Times[STATE-1])
    elif (5 == switch_1):
      $ 670 "Case 5"
      $ 671 "TM_St_Starting≔get_time(STATE_Times[STATE-1])"
      global TM_St_Starting=get_time(STATE_Times[STATE-1])
    elif (6 == switch_1):
      $ 672 "Case 6"
      $ 673 "TM_St_Execute≔get_time(STATE_Times[STATE-1])"
      global TM_St_Execute=get_time(STATE_Times[STATE-1])
    elif (7 == switch_1):
      $ 674 "Case 7"
      $ 675 "TM_St_Completin≔get_time(STATE_Times[STATE-1])"
      global TM_St_Completin=get_time(STATE_Times[STATE-1])
    elif (8 == switch_1):
      $ 676 "Case 8"
      $ 677 "TM_St_Complete≔get_time(STATE_Times[STATE-1])"
      global TM_St_Complete=get_time(STATE_Times[STATE-1])
    elif (9 == switch_1):
      $ 678 "Case 9"
      $ 679 "TM_St_Holding≔get_time(STATE_Times[STATE-1])"
      global TM_St_Holding=get_time(STATE_Times[STATE-1])
    elif (10 == switch_1):
      $ 680 "Case 10"
      $ 681 "TM_St_Held≔get_time(STATE_Times[STATE-1])"
      global TM_St_Held=get_time(STATE_Times[STATE-1])
    elif (11 == switch_1):
      $ 682 "Case 11"
      $ 683 "TM_St_Unholding≔get_time(STATE_Times[STATE-1])"
      global TM_St_Unholding=get_time(STATE_Times[STATE-1])
    elif (12 == switch_1):
      $ 684 "Case 12"
      $ 685 "TM_St_Suspendin≔get_time(STATE_Times[STATE-1])"
      global TM_St_Suspendin=get_time(STATE_Times[STATE-1])
    elif (13 == switch_1):
      $ 686 "Case 13"
      $ 687 "TM_St_Suspended≔get_time(STATE_Times[STATE-1])"
      global TM_St_Suspended=get_time(STATE_Times[STATE-1])
    elif (14 == switch_1):
      $ 688 "Case 14"
      $ 689 "TM_St_Unsuspend≔get_time(STATE_Times[STATE-1])"
      global TM_St_Unsuspend=get_time(STATE_Times[STATE-1])
    elif (15 == switch_1):
      $ 690 "Case 15"
      $ 691 "TM_St_Aborting≔get_time(STATE_Times[STATE-1])"
      global TM_St_Aborting=get_time(STATE_Times[STATE-1])
    elif (16 == switch_1):
      $ 692 "Case 16"
      $ 693 "TM_St_Aborted≔get_time(STATE_Times[STATE-1])"
      global TM_St_Aborted=get_time(STATE_Times[STATE-1])
    elif (17 == switch_1):
      $ 694 "Case 17"
      $ 695 "TM_St_Clearing≔get_time(STATE_Times[STATE-1])"
      global TM_St_Clearing=get_time(STATE_Times[STATE-1])
    end
    $ 697 "Wait: 0.1"
    sleep(0.1)
  end
end
